FUNCTION_BLOCK FB_HardwareOutputs
VAR_INPUT
    stOutputs : ST_HomeOutputs;
END_VAR


GVL_WorkshopIO.bLightRelay := stOutputs.Workshop.bLightRelay;
GVL_EntrywayIO.bLightRelay := stOutputs.Entryway.bLightRelay;
GVL_EntrywayIO.bTemporaryLightRelay := stOutputs.Entryway.bTemporaryLightRelay;
GVL_HallIO.bOuterSpotsRelay := stOutputs.Hall.bOuterSpotsRelay;
GVL_HallIO.bMiddleSpotRelay := stOutputs.Hall.bMiddleSpotRelay;

END_FUNCTION_BLOCK

(* stored: Version 1.1.0.1
   POU FB_HardwareOutputs: Id {734d95e1-63f5-4b5d-a283-35baa69a6c0e}, SpecialFunc None *)
